(* IEC 61131-3 sources: llm-plc-st-eval/data/definitivo/gpt-4o-2024-08-06/I2/zero_shot, 3 files *)

(* ---- ejec_1.st ---- *)
```pascal
FUNCTION_BLOCK FB_Llenado
VAR
    // Entradas
    nivelAlto : BOOL;
    nivelBajo : BOOL;
    btnInicio : BOOL;
    btnParo : BOOL;

    // Salidas
    vLlenado : BOOL := FALSE;
    motorMezcla : BOOL := FALSE;
    vDescarga : BOOL := FALSE;

    // Variables internas
    estado : INT := 0; // 0: Reposo, 1: Llenado, 2: Mezcla, 3: Descarga
    timerMezcla : TON; // Temporizador para la mezcla
END_VAR

// Inicialización del temporizador de mezcla
timerMezcla(IN := FALSE, PT := T#60S);

// Lógica de control del proceso
IF btnParo THEN
    // Si se presiona el botón de paro, se detiene el proceso y se desactivan todas las salidas
    estado := 0;
    vLlenado := FALSE;
    motorMezcla := FALSE;
    vDescarga := FALSE;
ELSE
    CASE estado OF
        0: // Estado de reposo
            IF btnInicio THEN
                estado := 1; // Iniciar llenado
            END_IF;

        1: // Estado de llenado
            vLlenado := TRUE;
            IF nivelAlto THEN
                vLlenado := FALSE;
                estado := 2; // Pasar a mezcla
                timerMezcla(IN := TRUE); // Iniciar temporizador de mezcla
            END_IF;

        2: // Estado de mezcla
            motorMezcla := TRUE;
            IF timerMezcla.Q THEN
                motorMezcla := FALSE;
                estado := 3; // Pasar a descarga
            END_IF;

        3: // Estado de descarga
            vDescarga := TRUE;
            IF nivelBajo THEN
                vDescarga := FALSE;
                estado := 0; // Volver a reposo
            END_IF;
    END_CASE;
END_IF;
END_FUNCTION_BLOCK
```

Este código implementa un proceso de llenado por etapas utilizando un bloque de función en Structured Text (ST) conforme al estándar IEC 61131-3. El proceso se controla mediante un estado interno que cambia en respuesta a las entradas y condiciones del sistema.

(* ---- ejec_2.st ---- *)
```pascal
FUNCTION_BLOCK FB_Llenado
VAR
    // Entradas
    nivelAlto : BOOL;   // Sensor de nivel alto
    nivelBajo : BOOL;   // Sensor de nivel bajo
    btnInicio : BOOL;   // Botón de inicio
    btnParo   : BOOL;   // Botón de paro

    // Salidas
    vLlenado   : BOOL;  // Válvula de llenado
    motorMezcla: BOOL;  // Motor de mezcla
    vDescarga  : BOOL;  // Válvula de descarga

    // Variables internas
    estadoProceso : INT;        // Estado del proceso
    timerMezcla   : TON;        // Temporizador para el motor de mezcla
END_VAR

// Inicialización
IF btnParo THEN
    // Si se presiona el botón de paro, reiniciar el proceso
    estadoProceso := 0;
    vLlenado := FALSE;
    motorMezcla := FALSE;
    vDescarga := FALSE;
ELSE
    CASE estadoProceso OF
        0: // Estado de reposo
            IF btnInicio THEN
                estadoProceso := 1; // Ir al estado de llenado
            END_IF;

        1: // Estado de llenado
            vLlenado := TRUE;
            IF nivelAlto THEN
                vLlenado := FALSE;
                estadoProceso := 2; // Ir al estado de mezcla
                timerMezcla(IN := TRUE, PT := T#60S); // Iniciar temporizador de mezcla
            END_IF;

        2: // Estado de mezcla
            motorMezcla := TRUE;
            timerMezcla(IN := TRUE);
            IF timerMezcla.Q THEN
                motorMezcla := FALSE;
                estadoProceso := 3; // Ir al estado de descarga
            END_IF;

        3: // Estado de descarga
            vDescarga := TRUE;
            IF nivelBajo THEN
                vDescarga := FALSE;
                estadoProceso := 0; // Volver al estado de reposo
            END_IF;
    END_CASE;
END_IF;
END_FUNCTION_BLOCK
```

Este código implementa un proceso de llenado por etapas en un bloque de función llamado `FB_Llenado`. El proceso se controla mediante un estado interno (`estadoProceso`) y responde a las entradas de los sensores y botones. El temporizador `timerMezcla` se utiliza para controlar el tiempo de operación del motor de mezcla.

(* ---- ejec_3.st ---- *)
```pascal
FUNCTION_BLOCK FB_Llenado
VAR_INPUT
    nivelAlto : BOOL;    // Sensor de nivel alto
    nivelBajo : BOOL;    // Sensor de nivel bajo
    btnInicio : BOOL;    // Botón de inicio
    btnParo   : BOOL;    // Botón de paro
END_VAR

VAR_OUTPUT
    vLlenado   : BOOL;   // Válvula de llenado
    motorMezcla: BOOL;   // Motor de mezcla
    vDescarga  : BOOL;   // Válvula de descarga
END_VAR

VAR
    estado     : INT;    // Estado del proceso
    timerMezcla: TON;    // Temporizador para el motor de mezcla
END_VAR

// Estados del proceso
// 0: Reposo
// 1: Llenado
// 2: Mezcla
// 3: Descarga

// Inicialización del bloque
IF NOT btnInicio THEN
    estado := 0;
END_IF

// Lógica de control del proceso
CASE estado OF
    0: // Reposo
        vLlenado := FALSE;
        motorMezcla := FALSE;
        vDescarga := FALSE;
        IF btnInicio THEN
            estado := 1;
        END_IF

    1: // Llenado
        vLlenado := TRUE;
        IF nivelAlto THEN
            vLlenado := FALSE;
            estado := 2;
            timerMezcla(IN := TRUE, PT := T#60S);
        END_IF

    2: // Mezcla
        motorMezcla := TRUE;
        timerMezcla(IN := TRUE);
        IF timerMezcla.Q THEN
            motorMezcla := FALSE;
            estado := 3;
        END_IF

    3: // Descarga
        vDescarga := TRUE;
        IF nivelBajo THEN
            vDescarga := FALSE;
            estado := 0;
        END_IF
END_CASE

// Lógica de paro de emergencia
IF btnParo THEN
    vLlenado := FALSE;
    motorMezcla := FALSE;
    vDescarga := FALSE;
    estado := 0;
END_IF

END_FUNCTION_BLOCK
```

Este código implementa un proceso de llenado por etapas utilizando el lenguaje Structured Text (ST) conforme al estándar IEC 61131-3. El proceso se controla mediante un bloque de función `FB_Llenado` que gestiona las entradas y salidas necesarias para el funcionamiento del sistema.
